(* IEC 61131-3 sources: trust-platform/manual-tests/root-a/src, 17 files *)

(* ---- InterfaceImpl.st ---- *)
INTERFACE IMotor
    METHOD Start : BOOL
    END_METHOD

    PROPERTY Speed : DINT
        GET
        END_GET
    END_PROPERTY
END_INTERFACE

CLASS Motor IMPLEMENTS IMotor
VAR
    speed : DINT;
END_VAR
END_CLASS

(* ---- MissingReturn.st ---- *)
FUNCTION MissingReturn : INT
VAR_INPUT
    a : INT;
END_VAR

(* missing return *)
END_FUNCTION

(* ---- NamespaceA.st ---- *)
NAMESPACE Core.Math
FUNCTION AddOne : DINT
VAR_INPUT
    X : DINT;
END_VAR
AddOne := X + 1;
END_FUNCTION
END_NAMESPACE

(* ---- NamespaceB.st ---- *)
NAMESPACE Vendor.LibA
FUNCTION AddOne : DINT
VAR_INPUT
    X : DINT;
END_VAR
AddOne := X + 10;
END_FUNCTION
END_NAMESPACE

(* ---- Main.st ---- *)
NAMESPACE Plant

CLASS Counter
VAR
    x : DINT;
END_VAR

PUBLIC METHOD Next : DINT
    x := x + 1;
    Next := x;
END_METHOD

PROPERTY Value : DINT
    GET
        Value := x;
    END_GET
END_PROPERTY

END_CLASS

FUNCTION AddTwo : DINT
VAR_INPUT
    A : DINT;
    B : DINT;
END_VAR
AddTwo := A + B;
END_FUNCTION

FUNCTION_BLOCK FB_Adder
VAR_INPUT
    A : DINT;
    B : DINT;
END_VAR
VAR_OUTPUT
    Result : DINT;
END_VAR
Result := A + B;
END_FUNCTION_BLOCK

PROGRAM Main
VAR
    counter : Counter;
    adder : FB_Adder;
    outVal : DINT;
    str : STRING;
    (* removed TIME and direct I/O for debug clarity *)
END_VAR

(* formal/non-formal mixing *)
outVal := AddTwo(1, 2);

(* formal before positional: reorder to positional-first *)
adder(2, 3, Result => outVal);

(* output binding operator fix *)
adder(A := 1, B := 2, Result => outVal);

(* simple literal assignment for debug *)
str := 'abc';

(* call hierarchy + refs *)
outVal := counter.Next();
END_PROGRAM

END_NAMESPACE

(* ---- Repro.st ---- *)
NAMESPACE Repro

INTERFACE IFoo
    METHOD Next : DINT
    END_METHOD
END_INTERFACE

CLASS Foo IMPLEMENTS IFoo
VAR
    x : DINT;
END_VAR

METHOD Next : DINT
    x := x + 1;
    Next := x;
END_METHOD
END_CLASS

FUNCTION AddTwo : DINT
VAR_INPUT
    A : DINT;
    B : DINT;
END_VAR
AddTwo := A + B;
END_FUNCTION

PROGRAM ReproMain
VAR
    foo : Foo;
    outVal : DINT;
END_VAR

outVal := AddTwo(A := 1, 2);
outVal := foo.Next();
END_PROGRAM

END_NAMESPACE

(* ---- Ambiguity.st ---- *)
USING Core.Math;
USING Vendor.LibA;

PROGRAM Ambiguity
VAR
    x : DINT;
END_VAR
x := AddOne(x); (* ambiguous; expect disambiguation quick fix *)
END_PROGRAM

(* ---- AmbiguityRepro.st ---- *)
USING Core.Math;
USING Vendor.LibA;

PROGRAM AmbiguityRepro
VAR
    x : DINT;
END_VAR
x := AddOne(x);
END_PROGRAM

(* ---- DebugMain.st ---- *)
PROGRAM DebugMain
VAR
    x : DINT := 1;
    y : DINT := 2;
    sum : DINT;
END_VAR

sum := x + y;
END_PROGRAM

(* ---- Formatting.st ---- *)
PROGRAM FormatTest
VAR
x:INT;
  y    :DINT;
END_VAR
x:=1; y :=2;(*comment*)
IF x=1 THEN
    y:=y+1;
END_IF
END_PROGRAM

(* ---- ImplicitConversion.st ---- *)
PROGRAM ImplicitConversion
VAR
    a : INT;
    b : BOOL;
END_VAR

b := a;
END_PROGRAM

(* ---- ImplicitConversion2.st ---- *)
PROGRAM ImplicitConversion2
VAR
    a : DINT;
    b : INT;
END_VAR

b := a;
END_PROGRAM

(* ---- MissingEndIf.st ---- *)
PROGRAM MissingEndIf
VAR
    a : INT;
END_VAR

IF a = 1 THEN
    a := 2;
END_IF
END_PROGRAM

(* ---- MissingType.st ---- *)
PROGRAM MissingType
VAR
    bad : MissingType;
END_VAR
END_PROGRAM

(* ---- MissingVar.st ---- *)
PROGRAM MissingVar
VAR
    a : INT;
END_VAR

b := a;
END_PROGRAM

(* ---- Tasks.st ---- *)
CONFIGURATION PlantConfig
RESOURCE Res1 ON PLC
    TASK FastTask(INTERVAL := T#10ms, PRIORITY := 1);
    TASK SlowTask(INTERVAL := T#100ms, PRIORITY := 10);

    PROGRAM P1 WITH FastTask : Main;
    PROGRAM P2 WITH SlowTask : Main;
END_RESOURCE
END_CONFIGURATION

(* ---- TasksBad.st ---- *)
CONFIGURATION BadConfig
RESOURCE Res1 ON PLC
    TASK BadTask(INTERVAL := T#10ms);
END_RESOURCE
END_CONFIGURATION
